// TIA Portal V19 export
VAR_GLOBAL   // PLC tag table "Default tag table"
   Axis_1_Drive_IN AT %I68.0 : "PD_TEL3_IN";
   Axis_1_Drive_OUT AT %Q64.0 : "PD_TEL3_OUT";
   HSC_1_Up AT %I0.0 : Bool;
   HSC_1_Down AT %I0.1 : Bool;
   Tag_1 AT %ID78 : DInt;
   Tag_2 AT %ID82 : DWord;
END_VAR
VAR_GLOBAL CONSTANT   // user constants
   INV_CMD_FORW : Word := 16#0031;
   INV_CMD_STOP : Word := 16#0022;
   INV_CMD_REV : Word := 16#0032;   // !!! CHECK
   TYPE_CONV_1 : Int := 2;
   TYPE_CONV_2 : Int := 1;
   CONV_1_DRUM_DIA : Real := 82.0;   // mm
   CONV_1_MOTOR_RPM : Real := 1365.0;
   CONV_1_REDUCER_I : Real := 10.0;
   C1_CONV_ID : Int := 1;
   CONV_2_PITCH : Real := 33.0;   // mm
   CONV_2_MOTOR_RPM : Real := 1365.0;   // Nominal RPM at 50 Hz
   C2_CONV_ID : Int := 2;
   PI : Real := 3.14159265358;
   CONV_2_DRUM_Z : Real := 14.0;
   CONV_2_REDUCER_I : Real := 30.0;
   ROBOT_CMD_APPROACH_PICK : Int := 20;
   ROBOT_CMD_GO_HOME : Int := 10;
   ROBOT_CMD_PICK : Int := 30;
   ROBOT_CMD_APPROACH_PLACE : Int := 40;
   ROBOT_CMD_PLACE : Int := 50;
END_VAR
